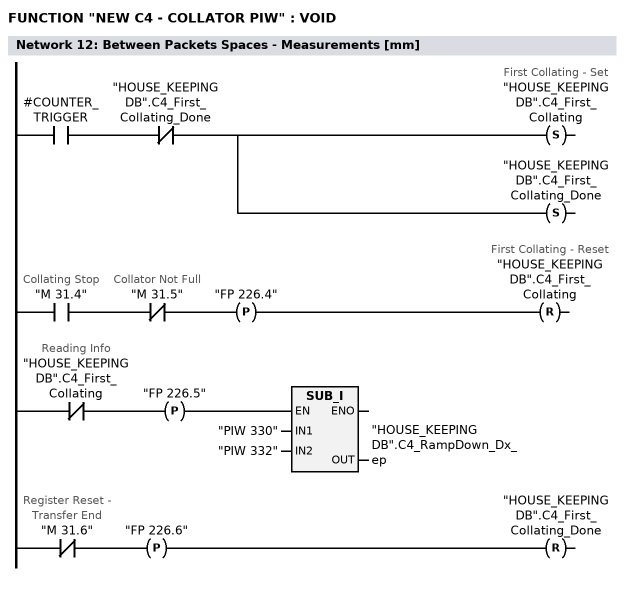

      A     #COUNTER_TRIGGER;
      AN    "HOUSE_KEEPING DB".C4_First_Collating_Done;
      S     "HOUSE_KEEPING DB".C4_First_Collating; // First Collating - Set
      S     "HOUSE_KEEPING DB".C4_First_Collating_Done;
//;
      A     "M 31.4"; // Collating Stop
      AN    "M 31.5"; // Collator Not Full
      FP    "FP 226.4";
      R     "HOUSE_KEEPING DB".C4_First_Collating; // First Collating - Reset
//;
      AN    "HOUSE_KEEPING DB".C4_First_Collating; // Reading Info
      FP    "FP 226.5";
      JCN   N1ST;

      L     "PIW 330"; // Direct Ch3 (was ACT_CNTV3, ~100 mS old)
      L     "PIW 332"; // Direct Ch2 (was ACT_CNTV2, ~100 mS old)
      -I    ;
      T     "HOUSE_KEEPING DB".C4_RampDown_Dx_ep;

N1ST: NOP   0;

      AN    "M 31.6"; // Register Reset - Transfer End
      FP    "FP 226.6";
      R     "HOUSE_KEEPING DB".C4_First_Collating_Done;
NETWORK
TITLE =Conveyor 4 - Surface Length Left (PulseUnit) - Measurements

      A     "M 31.1";
      S     "M 166.3";
//;
      A     "M 166.3";
      AN    "M 31.7";
      =     "FM350 DB".CONTROL_SIGNALS.SW_GATE3;
//;
      A     "M 166.3";
      A     "M 31.1";
      JNB   M663;
      L     "COLLATORS DB".Surface_Length_C4;
      L     "PIW 330"; // Direct Ch3 (was ACT_CNTV3, ~100 mS old)
      -D    ;
      T     "COLLATORS DB".Surface_Left_C4;
      L     0;
      >=I   ;
      JNB   T004;
      L     "COLLATORS DB".Surface_Left_C4;
      T     "COLLATORS DB".Surface_Length_Left_C4;

T004: CLR   ;

M663: CLR   ;
NETWORK
TITLE =Conveyor 4 - Space Between - Calculator

      A     "M 167.1";
      FP    "FP 154.2";
      JNB   M581;
      L     "COLLATORS DB".Surface_Left_C4;
      L     "COLLATORS DB".Frac_Packet_Length_C4;
      -I    ;
      T     "MW 214";

M581: CLR   ;

      A     "M 167.1";
      JNB   M671;
      A(    ;
      L     "COLLATORS DB".Surface_Left_C4;
      L     "MW 214";
      <=I   ;
      )     ;
      R     "M 167.1";

M671: CLR   ;
NETWORK
TITLE =Conveyor 4 - Collating Length Manager

      A     "M 166.3";
      AN    "M 30.4";
      A     "M 31.4";
      JNB   M304;
      L     "COLLATORS DB".Surface_Left_C4;
      L     "COLLATORS DB".Packet_Length_Frac_C4;
      <I    ;
      S     "M 30.4";

M304: CLR   ;

      A     "M 10.1";
      FP    "FP 154.7";
      O     "M 31.7";
      R     "M 30.4";
NETWORK
TITLE =Packet Length to HMI + Hysteresis

      A     "M 167.4";
      JNB   C167;
      A(    ;
      A(    ;
      L     "MW 202";
      L     "MW 204";
      >I    ;
      )     ;
      O     ;
      A(    ;
      L     "MW 202";
      L     "MW 206";
      <I    ;
      )     ;
      )     ;
      JNB   BYP5;
      L     "MW 202";
      T     "HMI_DB".WORD_PACKET_LENGTH;

BYP5: CLR   ;

      L     "MW 202";
      L     3.000000e+000;
      *R    ;
      L     1.000000e+002;
      /R    ;
      T     #R_TUBE_PERCENT;
      TRUNC ;
      T     #W_TUBE_PERCENT;
//;
      L     #W_TUBE_PERCENT;
      L     "MW 202";
      +I    ;
      T     "MW 204";
//;
      L     #W_TUBE_PERCENT;
      L     "MW 202";
      -I    ;
      T     "MW 206";
//;
      CLR   ;
      =     "M 167.4";

C167: CLR   ;
NETWORK
TITLE =Collator
//Collator House Keeping


NETWORK
TITLE =Collator Conveyor 4 - Clearing
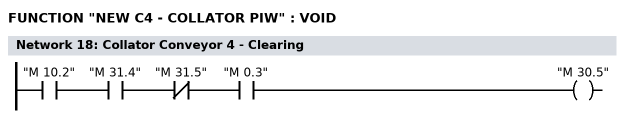

      A     "M 10.2";
      A     "M 31.4";
      AN    "M 31.5";
      A     "M 0.3";
      =     "M 30.5";
NETWORK
TITLE =Soft Timer 33 Reset - Clearing TimeOut 20s + Freeze Option

      A     "M 30.5";
      A     "A 44.3";
      A     "M 0.3";
      JCN   R331;
      JU    E331;

R331: L     L#0;
      T     "DB UTILITY".T33_ET;
      R     "DB UTILITY".T33_DN;

E331: NOP   0;
NETWORK
TITLE =Soft Timer 33 Add

      A     "M 30.5";
      A     "A 44.3";
      A     "M 0.3";
      AN    "DB UTILITY".Freeze_Sequence_2;
      AN    "DB UTILITY".T33_DN;
      JCN   E332;

      L     "DB UTILITY".T33_ET;
      L     "DB UTILITY".Scan_Cycle_Previous;
      ITD   ;
      +D    ;
      T     "DB UTILITY".T33_ET;

E332: NOP   0;
NETWORK
TITLE =Soft Timer 33 Done 20s

      L     "DB UTILITY".T33_ET;
      L     L#20000;
      >=D   ;
      =     "DB UTILITY".T33_DN;
NETWORK
TITLE =Collator Conveyor 4 - Clearing Surface - Run 2K Encoder Counts

      A     "M 30.5";
      A     "A 44.3";
      A     "M 0.3";
      JNB   M305;
      A(    ;
      L     "PIW 332"; // Direct Ch2 (was ACT_CNTV2, ~100 mS old)
      L     2000;
      >I    ;
      )     ;
      =     "M 30.3";

M305: CLR   ;
NETWORK
TITLE =Collator Conveyor 4 - Packet at the End !
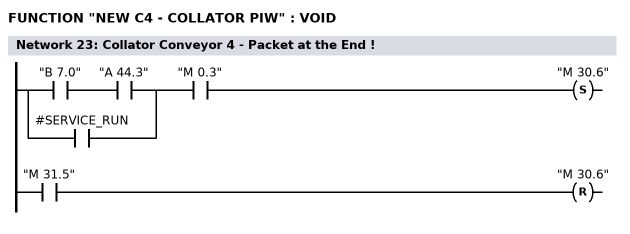

      A     "B 7.0";
      A     "A 44.3";
      O     #SERVICE_RUN;
      A     "M 0.3";
      S     "M 30.6";
//;
      A     "M 31.5";
      R     "M 30.6";
NETWORK
TITLE =Soft Timer 31 Reset - InFeed TimeOut 5s With Freeze Option

      A     "M 31.2";
      AN    "M 31.4";
      A     "A 44.3";
      A     "M 0.3";
      JCN   R311;
      JU    E311;

R311: L     L#0;
      T     "DB UTILITY".T31_ET;
      R     "DB UTILITY".T31_DN;

E311: NOP   0;
NETWORK
TITLE =Soft Timer 31 Add

      A     "M 31.2";
      AN    "M 31.4";
      A     "A 44.3";
      A     "M 0.3";
      AN    "DB UTILITY".Freeze_Sequence_2;
      AN    "DB UTILITY".T31_DN;
      JCN   E312;

      L     "DB UTILITY".T31_ET;
      L     "DB UTILITY".Scan_Cycle_Previous;
      ITD   ;
      +D    ;
      T     "DB UTILITY".T31_ET;

E312: NOP   0;
NETWORK
TITLE =Soft Timer 31 Done 5s
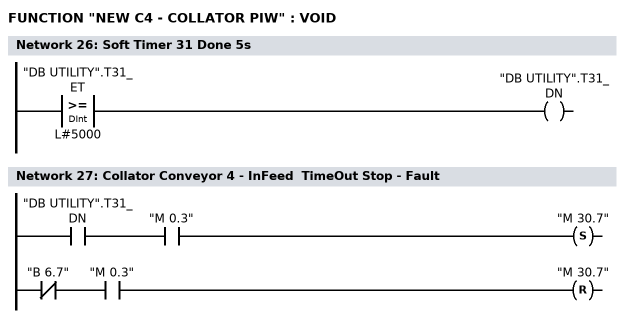

      L     "DB UTILITY".T31_ET;
      L     L#5000;
      >=D   ;
      =     "DB UTILITY".T31_DN;
NETWORK
TITLE =Collator Conveyor 4 - InFeed  TimeOut Stop - Fault

      A     "DB UTILITY".T31_DN;
      A     "M 0.3";
      S     "M 30.7";
//;
      AN    "B 6.7";
      A     "M 0.3";
      R     "M 30.7";
NETWORK
TITLE =Collator
//Collator Steps


NETWORK
TITLE =Collator Conveyor 4 - Steps Register - Reset

      A(    ;
      O     "M 31.7";
      O     "DB UTILITY".T33_DN;
      O     #INITIALISATION;
      O     "DB UTILITY".Conveyor_4_Disable;
      )     ;
      A     "M 0.3";
      JNB   INIT;
      L     W#16#0;
      T     "MW 31";
      S     "M 167.0";

INIT: CLR   ;
NETWORK
TITLE =Step 5N1  - Power ON
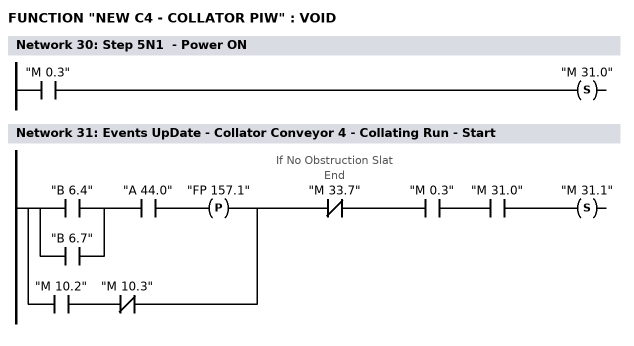

      A     "M 0.3";
      S     "M 31.0";
NETWORK
TITLE =Events UpDate - Collator Conveyor 4 - Collating Run - Start

      A(    ;
      A(    ;
      O     "B 6.4";
      O     "B 6.7";
      )     ;
      A     "A 44.0";
      FP    "FP 157.1";
      O     ;
      A     "M 10.2";
      AN    "M 10.3";
      )     ;
      AN    "M 33.7"; // If No Obstruction Slat End
      A     "M 0.3";
      A     "M 31.0";
      S     "M 31.1";
NETWORK
TITLE =Soft Timer 29 Reset - LB Obstruction Alarm 10s + Freeze Option

      A(    ;
      O     "B 6.4";
      O     "B 6.7";
      )     ;
      AN    "A 44.0";
      JCN   R281;
      JU    E281;

R281: L     L#0;
      T     "DB UTILITY".T29_ET;
      R     "DB UTILITY".T29_DN;

E281: NOP   0;
NETWORK
TITLE =Soft Timer 29 Add

      A(    ;
      O     "B 6.4";
      O     "B 6.7";
      )     ;
      AN    "A 44.0";
      AN    "DB UTILITY".Freeze_Sequence_2;
      AN    "DB UTILITY".T29_DN;
      JCN   E282;

      L     "DB UTILITY".T29_ET;
      L     "DB UTILITY".Scan_Cycle_Previous;
      ITD   ;
      +D    ;
      T     "DB UTILITY".T29_ET;

E282: NOP   0;
NETWORK
TITLE =Soft Timer 29 Done 10s
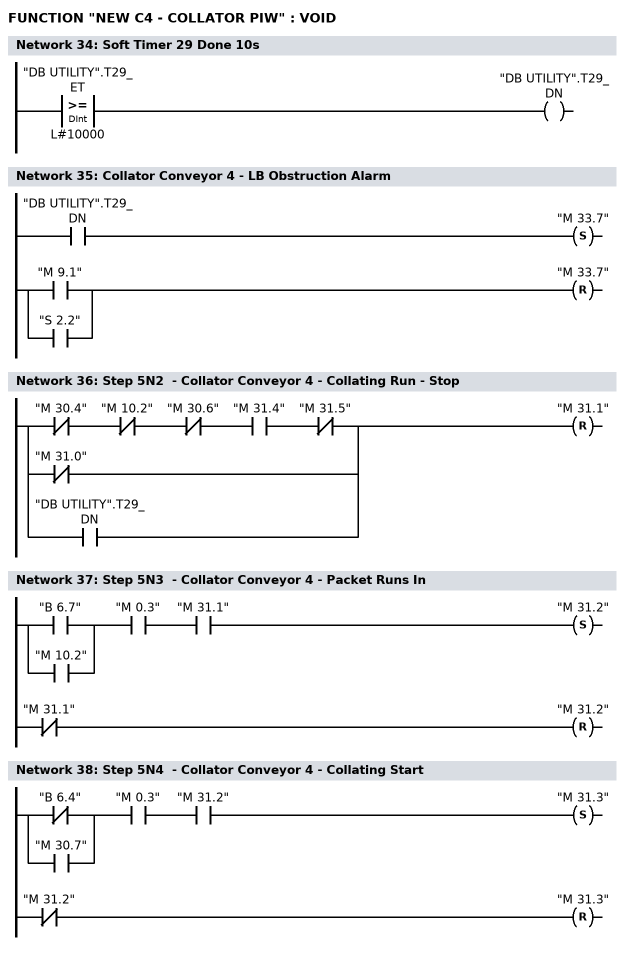

      L     "DB UTILITY".T29_ET;
      L     L#10000;
      >=D   ;
      =     "DB UTILITY".T29_DN;
NETWORK
TITLE =Collator Conveyor 4 - LB Obstruction Alarm

      A     "DB UTILITY".T29_DN;
      S     "M 33.7";
//;
      A(    ;
      O     "M 9.1";
      O     "S 2.2";
      )     ;
      R     "M 33.7";
NETWORK
TITLE =Step 5N2  - Collator Conveyor 4 - Collating Run - Stop

      A(    ;
      AN    "M 30.4";
      AN    "M 10.2";
      AN    "M 30.6";
      A     "M 31.4";
      AN    "M 31.5";
      ON    "M 31.0";
      O     "DB UTILITY".T29_DN;
      )     ;
      R     "M 31.1";
NETWORK
TITLE =Step 5N3  - Collator Conveyor 4 - Packet Runs In

      A(    ;
      O     "B 6.7";
      O     "M 10.2";
      )     ;
      A     "M 0.3";
      A     "M 31.1";
      S     "M 31.2";
//;
      AN    "M 31.1";
      R     "M 31.2";
NETWORK
TITLE =Step 5N4  - Collator Conveyor 4 - Collating Start

      A(    ;
      ON    "B 6.4";
      O     "M 30.7";
      )     ;
      A     "M 0.3";
      A     "M 31.2";
      S     "M 31.3";
//;
      AN    "M 31.2";
      R     "M 31.3";
NETWORK
TITLE =Step 5N5  - Collator Conveyor 4 - Collating Stop

      A(    ;
      AN    "B 6.7";
      AN(   ;
      AN    "M 10.2";
      A     "M 167.1";
      )     ;
      O     "M 30.7";
      )     ;
      A     "M 0.3";
      A     "M 31.3";
      S     "M 31.4";
//;
      AN    "M 31.3";
      R     "M 31.4";
NETWORK
TITLE =Step 5N6  - Collator Conveyor 4 - Full - Start Transfer
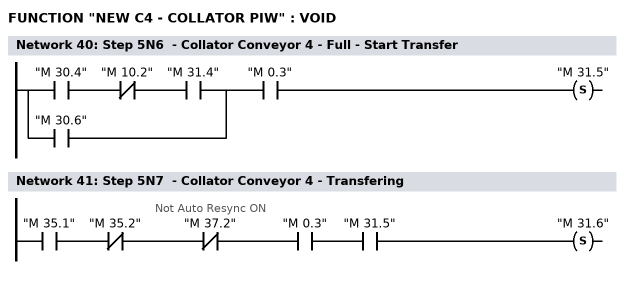

      A(    ;
      A     "M 30.4";
      AN    "M 10.2";
      A     "M 31.4";
      O     "M 30.6";
      )     ;
      A     "M 0.3";
      S     "M 31.5";
NETWORK
TITLE =Step 5N7  - Collator Conveyor 4 - Transfering

      A     "M 35.1";
      AN    "M 35.2";
      AN    "M 37.2"; // Not Auto Resync ON
      A     "M 0.3";
      A     "M 31.5";
      S     "M 31.6";
NETWORK
TITLE =Soft Timer 32 Reset - Transfer TimeOut 20s + Freeze Option

      A     "M 31.6";
      AN    "M 31.7";
      A     "A 44.3";
      A     "M 0.3";
      JCN   R321;
      JU    E321;

R321: L     L#0;
      T     "DB UTILITY".T32_ET;
      R     "DB UTILITY".T32_DN;

E321: NOP   0;
NETWORK
TITLE =Soft Timer 32 Add

      A     "M 31.6";
      AN    "M 31.7";
      A     "A 44.3";
      A     "M 0.3";
      AN    "DB UTILITY".Freeze_Sequence_2;
      AN    "DB UTILITY".T32_DN;
      JCN   E322;

      L     "DB UTILITY".T32_ET;
      L     "DB UTILITY".Scan_Cycle_Previous;
      ITD   ;
      +D    ;
      T     "DB UTILITY".T32_ET;

E322: NOP   0;
NETWORK
TITLE =Soft Timer 32 Done 20s
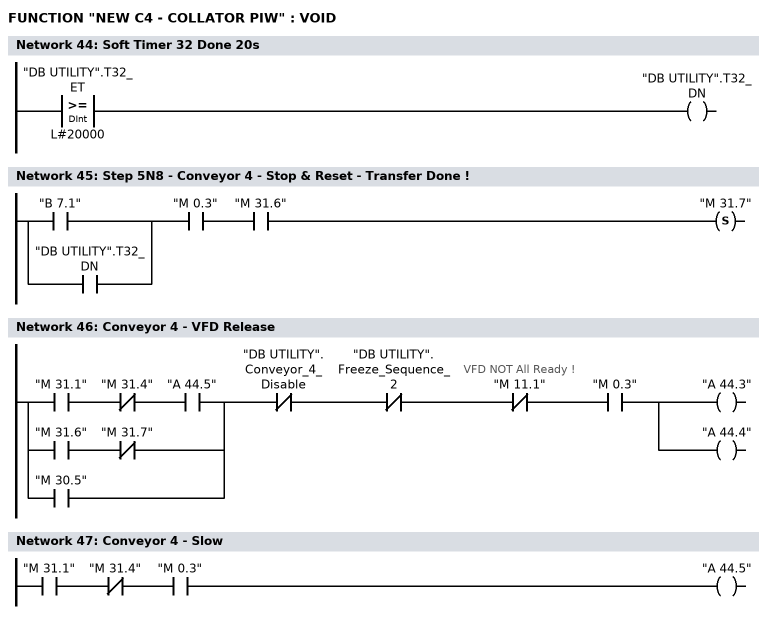

      L     "DB UTILITY".T32_ET;
      L     L#20000;
      >=D   ;
      =     "DB UTILITY".T32_DN;
NETWORK
TITLE =Step 5N8 - Conveyor 4 - Stop & Reset - Transfer Done !

      A(    ;
      O     "B 7.1";
      O     "DB UTILITY".T32_DN;
      )     ;
      A     "M 0.3";
      A     "M 31.6";
      S     "M 31.7";
NETWORK
TITLE =Conveyor 4 - VFD Release

      A(    ;
      A     "M 31.1";
      AN    "M 31.4";
      A     "A 44.5";
      O     ;
      A     "M 31.6";
      AN    "M 31.7";
      O     "M 30.5";
      )     ;
      AN    "DB UTILITY".Conveyor_4_Disable;
      AN    "DB UTILITY".Freeze_Sequence_2;
      AN    "M 11.1"; // VFD NOT All Ready !
      A     "M 0.3";
      =     "A 44.3";
      =     "A 44.4";
NETWORK
TITLE =Conveyor 4 - Slow

      A     "M 31.1";
      AN    "M 31.4";
      A     "M 0.3";
      =     "A 44.5";
END_FUNCTION

FUNCTION "NEW C5 - LINK" : VOID
TITLE =NEW FC934 (was FC1034) - Conveyor 5 - Link Pos.7
//Using "Soft Timer" cause S5T Timer cannot Pause/Freeze !...
NAME : POS_7
VERSION : 0.0


VAR_TEMP
  MAIN_SERVICE_2_SW : BOOL ;
  SERVICE_RUN : BOOL ;
  INITIALISATION : BOOL ;
END_VAR
BEGIN
NETWORK
TITLE =Conveyor 5 - Service

      A     "HMI_DB".ALL_SERVICE_ENABLE_SW;
      A     "HMI_DB".CONVEYOR_5_SERVICE_SW;
      A     "HMI_DB".SERVICE_SW_2_STATUS;
      =     #MAIN_SERVICE_2_SW;
//;
      A     #MAIN_SERVICE_2_SW;
      O     "M 34.1";
      JNB   CON5;
//;
      A     "HMI_DB".HMI_CONVEYOR_5_TEST_SSW;
      AN    "A 44.3";
      =     #SERVICE_RUN;
      S     "DB UTILITY".Conveyor_4_Disable;
//;
      A     "HMI_DB".SERVICE_INIT_PB;
      =     #INITIALISATION;
//;
      AN    #MAIN_SERVICE_2_SW;
      R     "HMI_DB".HMI_CONVEYOR_5_TEST_SSW;
      R     "DB UTILITY".Conveyor_4_Disable;

CON5: R     #SERVICE_RUN;
      R     #INITIALISATION;
      FP    "FP 158.5";
      =     "M 34.1";

NETWORK
TITLE =Service Mode
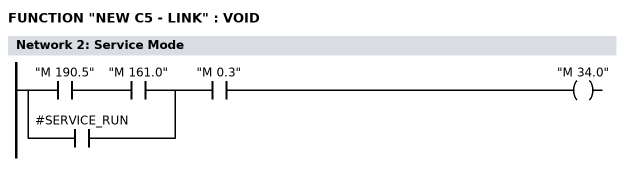

      A(    ;
      A     "M 190.5";
      A     "M 161.0";
      O     ;
      A     #SERVICE_RUN;
      )     ;
      A     "M 0.3";
      =     "M 34.0";

NETWORK
TITLE =Conveyor 5 - Steps Register - Reset

      A(    ;
      A     "M 35.1";
      AN    "M 35.2";
      A     "DB UTILITY".T35_DN;
      O     "M 35.4";
      O     #INITIALISATION;
      O     "DB UTILITY".Conveyor_5_Disable;
      )     ;
      A     "M 0.3";
      JC    M001;
      JU    M002;

M001: L     W#16#0;
      T     "MW 35";
      T     "HMI DB NEW".CONV_5_COUNT;

M002: NOP   0;

NETWORK
TITLE =Step 6N1 - Power ON
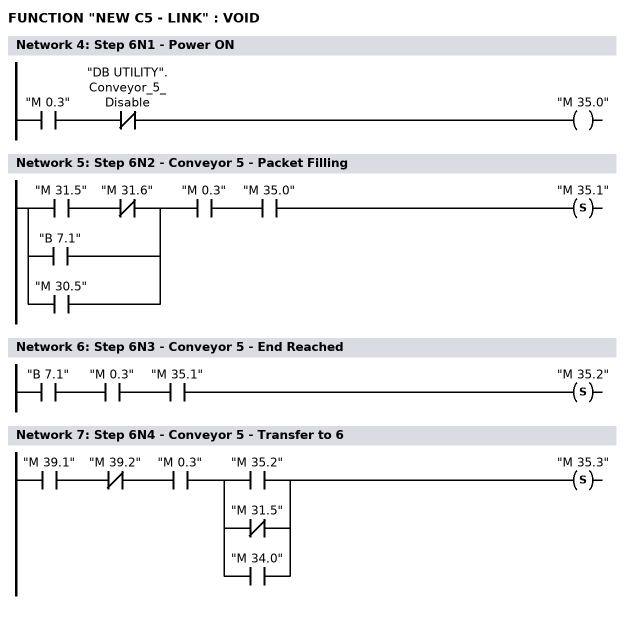

      A     "M 0.3";
      AN    "DB UTILITY".Conveyor_5_Disable;
      =     "M 35.0";

NETWORK
TITLE =Step 6N2 - Conveyor 5 - Packet Filling

      A(    ;
      A     "M 31.5";
      AN    "M 31.6";
      O     "B 7.1";
      O     "M 30.5";
      )     ;
      A     "M 0.3";
      A     "M 35.0";
      S     "M 35.1";

NETWORK
TITLE =Step 6N3 - Conveyor 5 - End Reached

      A     "B 7.1";
      A     "M 0.3";
      A     "M 35.1";
      S     "M 35.2";

NETWORK
TITLE =Step 6N4 - Conveyor 5 - Transfer to 6

      A     "M 39.1";
      AN    "M 39.2";
      A     "M 0.3";
      A(    ;
      O     "M 35.2";
      ON    "M 31.5";
      O     "M 34.0";
      )     ;
      S     "M 35.3";

NETWORK
TITLE =Soft Timer 35 Reset

      A(    ;
      A     "M 35.1";
      AN    "M 35.2";
      O     ;
      A     "M 35.3";
      AN    "M 35.4";
      A     "A 45.0";
      )     ;
      A     "M 0.3";
      JCN   R351;
      JU    E351;

R351: L     L#0;
      T     "DB UTILITY".T35_ET;
      R     "DB UTILITY".T35_DN;

E351: NOP   0;

NETWORK
TITLE =Soft Timer 35 Add

      A(    ;
      A     "M 35.1";
      AN    "M 35.2";
      O     ;
      A     "M 35.3";
      AN    "M 35.4";
      A     "A 45.0";
      )     ;
      A     "M 0.3";
      JCN   E352;
//;
      A     "DB UTILITY".Freeze_Sequence_2;
      A     "M 35.1";
      AN    "M 35.2";
      JC    E352;
//;
      AN    "DB UTILITY".T35_DN;
      JCN   E352;
//;
      L     "DB UTILITY".T35_ET;
      L     "DB UTILITY".Scan_Cycle_Previous;
      ITD   ;
      +D    ;
      T     "DB UTILITY".T35_ET;

E352: NOP   0;

NETWORK
TITLE =Soft Timer 35 Done 30s

      L     "DB UTILITY".T35_ET;
      L     L#30000; // [mS]
      >=D   ;
      =     "DB UTILITY".T35_DN;

NETWORK
TITLE =Automatic Re-Synchronization
//In Order to keep Synchronized,
//if Every Conditions are there, Conveyor 5 will do a Synchro Run 13sec after
//every 5 runs !
      A     "A 45.0"; // Count runs
      FP    "FP 169.7";
      JNB   ARS1;

      L     "MW 220"; // Count up
      L     1;
      +I    ;
      T     "MW 220";
//;
      L     10;
      >=I   ;
      JNB   ARS1;
//;
      S     "M 37.3"; // ARM after 5 runs
      L     0;
      T     "MW 220";

ARS1: NOP   0;

      A     "M 37.3"; // ARMED
      AN    "M 37.2"; // NOT already running
      AN    "DB UTILITY".Freeze_Sequence_2;
      AN    "A 45.0"; // wait end of run
      A     "M 35.0"; // power ON
      AN    "M 35.4"; // not in reset/stop
      JNB   ARS2;
//;
      L     "HMI_DB".CONV_4_COUNT; // Conveyor 4 Must be <= 2
      L     3;
      <I    ;
      JNB   ARS2;
//;
      L     "HMI_DB".CONV_5_COUNT;
      L     0; // Conveyor 5 Must NOT be Empty
      >I    ;
      JNB   ARS2;
//;
      L     "HMI_DB".CONV_6_COUNT;
      L     0; // Conveyor 6 Must be Empty
      ==I   ;
      JNB   ARS2;
//;
      AN    "B 7.2"; // Conveyor 6 Must be Empty
      AN    "M 10.0"; // Not Clearing
      JNB   ARS2;
//;
      S     "M 37.2"; // START 13s RUN
      R     "M 37.3"; // DISARM

ARS2: NOP   0;

      A     "M 37.2"; // Re-Sync ON
      L     S5T#13S;
      SD    "Timer 64";
//;
      A     "Timer 64"; // End Re-Sync if TimeOut 13s
      O     "B 7.1"; // or if Packet at END Sensor
      R     "M 37.2"; // Re-Sync OFF
NETWORK
TITLE =Automatic Re-Synchronization - Arm Timeout
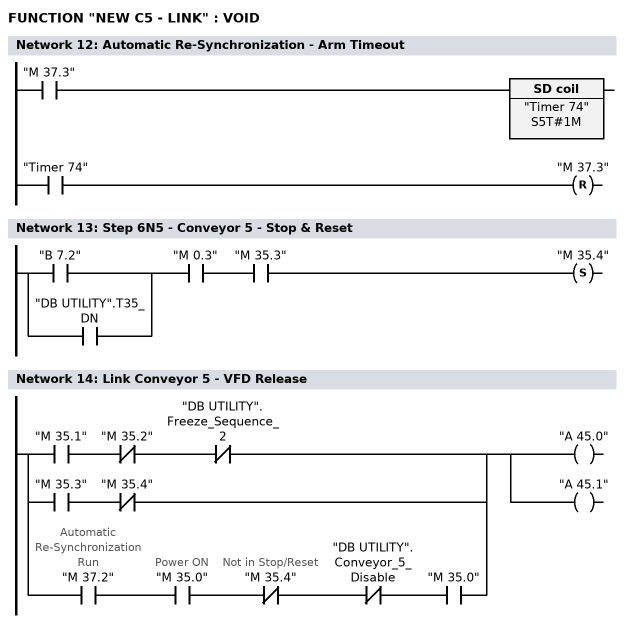

      A     "M 37.3";
      L     S5T#1M;
      SD    "Timer 74";
//;
      A     "Timer 74";
      R     "M 37.3";
NETWORK
TITLE =Step 6N5 - Conveyor 5 - Stop & Reset

      A(    ;
      O     "B 7.2";
      O     "DB UTILITY".T35_DN;
      )     ;
      A     "M 0.3";
      A     "M 35.3";
      S     "M 35.4";

NETWORK
TITLE =Link Conveyor 5 - VFD Release

      A(    ;
      A(    ;
      A     "M 35.1";
      AN    "M 35.2";
      AN    "DB UTILITY".Freeze_Sequence_2;
      )     ;
      O     ;
      A     "M 35.3";
      AN    "M 35.4";
      )     ;
      O     ;
      A(    ;
      A     "M 37.2"; // Automatic Re-Synchronization Run
      A     "M 35.0"; // Power ON
      AN    "M 35.4"; // Not in Stop/Reset
      )     ;
      AN    "DB UTILITY".Conveyor_5_Disable;
      A     "M 35.0";
      =     "A 45.0";
      =     "A 45.1";
END_FUNCTION

FUNCTION "NEW C6 - FLIP DELIV." : VOID
TITLE =NEW FC938 (was FC1038) - Conveyor 6 - Delivery to Flipper Pos.8
NAME : POS_8
VERSION : 0.0


VAR_TEMP
  MAIN_SERVICE_2_SW : BOOL ;
  SERVICE_RUN : BOOL ;
  INITIALISATION : BOOL ;
END_VAR
BEGIN
NETWORK
TITLE =Slat Conveyor - Service

      A     "HMI_DB".ALL_SERVICE_ENABLE_SW;
      A     "HMI_DB".CONVEYOR_6_SERVICE_SW;
      A     "HMI_DB".SERVICE_SW_2_STATUS;
      =     #MAIN_SERVICE_2_SW;
      CLR   ; // Fix: #INITIALISATION was never written
      =     #INITIALISATION;
//;
      A     #MAIN_SERVICE_2_SW;
      O     "M 38.1";
      JNB   CON6;
      A     "HMI_DB".HMI_CONVEYOR_6_TEST_SSW;
      =     #SERVICE_RUN;
      S     "DB UTILITY".Conveyor_5_Disable;
//;
      AN    #MAIN_SERVICE_2_SW;
      R     "HMI_DB".HMI_CONVEYOR_6_TEST_SSW;
      R     "DB UTILITY".Conveyor_5_Disable;

CON6: R     #SERVICE_RUN;
      R     #INITIALISATION;
      FP    "FP 158.6";
      =     "M 38.1";
NETWORK
TITLE =Flipper Delivery Conveyor 6 - Running TimeOut  30s
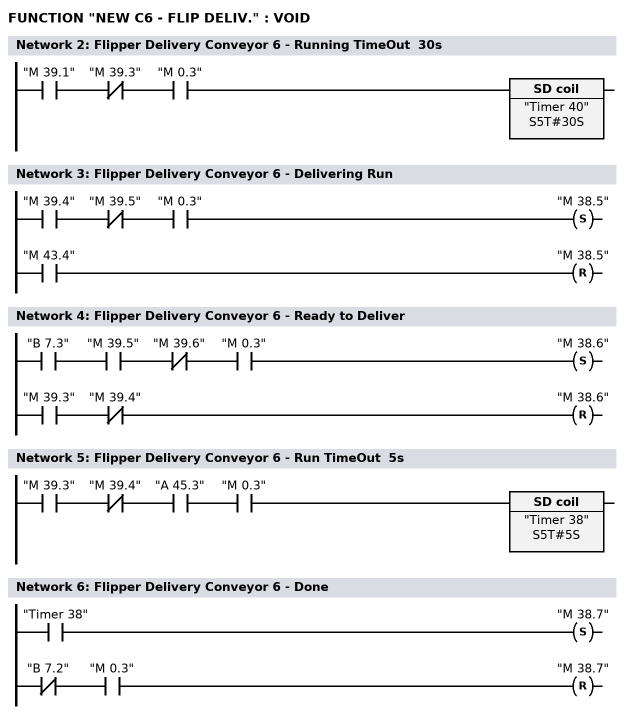

      A     "M 39.1";
      AN    "M 39.3";
      A     "M 0.3";
      L     S5T#30S;
      SD    "Timer 40";
NETWORK
TITLE =Flipper Delivery Conveyor 6 - Delivering Run

      A     "M 39.4";
      AN    "M 39.5";
      A     "M 0.3";
      S     "M 38.5";
//;
      A     "M 43.4";
      R     "M 38.5";
NETWORK
TITLE =Flipper Delivery Conveyor 6 - Ready to Deliver

      A     "B 7.3";
      A     "M 39.5";
      AN    "M 39.6";
      A     "M 0.3";
      S     "M 38.6";
//;
      A     "M 39.3";
      AN    "M 39.4";
      R     "M 38.6";
NETWORK
TITLE =Flipper Delivery Conveyor 6 - Run TimeOut  5s

      A     "M 39.3";
      AN    "M 39.4";
      A     "A 45.3";
      A     "M 0.3";
      L     S5T#5S;
      SD    "Timer 38";
NETWORK
TITLE =Flipper Delivery Conveyor 6 - Done

      A     "Timer 38";
      S     "M 38.7";
//;
      AN    "B 7.2";
      A     "M 0.3";
      R     "M 38.7";
NETWORK
TITLE =Conveyor 6 - Steps Register - Reset

      A(    ;
      O     "M 39.6";
      O     "Timer 40";
      O     #INITIALISATION;
      O     "DB UTILITY".Conveyor_6_Disable;
      )     ;
      A     "M 0.3";
      JC    M001;
      JU    M002;

M001: L     W#16#0;
      T     "MW 39";
      T     "MB 41";
      T     "HMI DB NEW".CONV_6_COUNT;

M002: NOP   0;
NETWORK
TITLE =Step 7N1 - Power ON
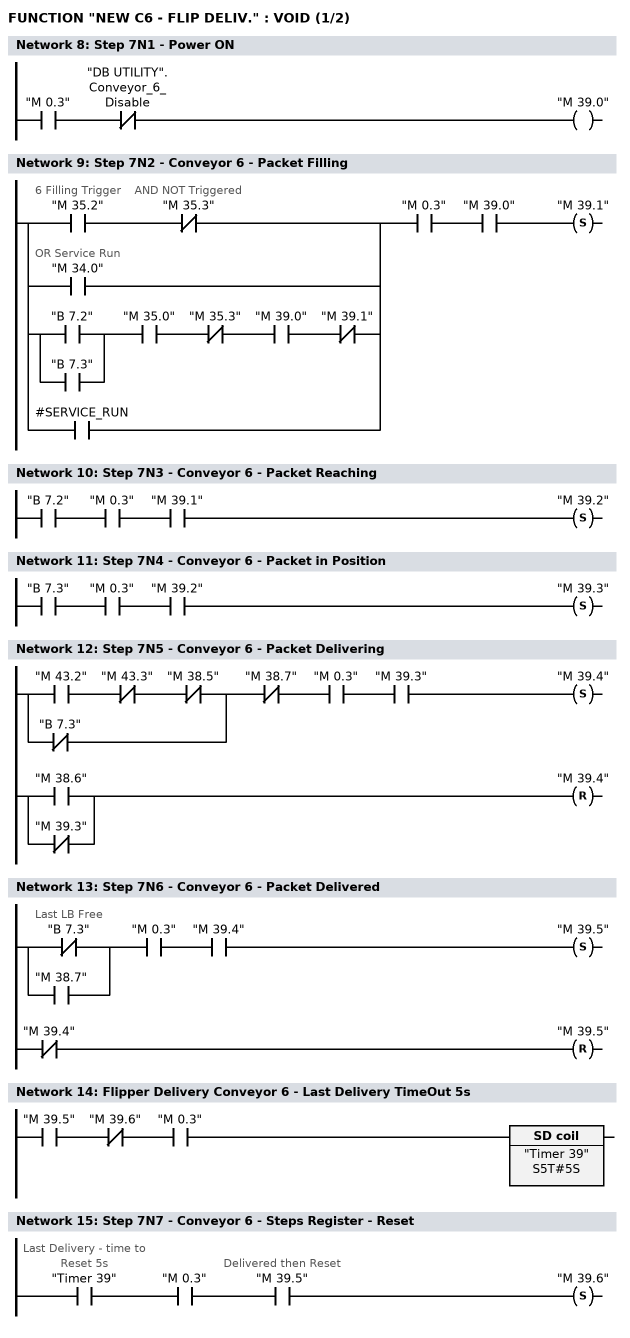

      A     "M 0.3";
      AN    "DB UTILITY".Conveyor_6_Disable;
      =     "M 39.0";
NETWORK
TITLE =Step 7N2 - Conveyor 6 - Packet Filling

      A(    ;

      A     "M 35.2"; // 6 Filling Trigger
      AN    "M 35.3"; // AND NOT Triggered
      O     "M 34.0"; // OR Service Run

      O     ;

      A(    ;
      O     "B 7.2";
      O     "B 7.3";
      )     ;
      A     "M 35.0";
      AN    "M 35.3";
      A     "M 39.0";
      AN    "M 39.1";

      O     ;

      A     #SERVICE_RUN;
      )     ;

      A     "M 0.3";
      A     "M 39.0";
      S     "M 39.1";
NETWORK
TITLE =Step 7N3 - Conveyor 6 - Packet Reaching

      A     "B 7.2";
      A     "M 0.3";
      A     "M 39.1";
      S     "M 39.2";
NETWORK
TITLE =Step 7N4 - Conveyor 6 - Packet in Position

      A     "B 7.3";
      A     "M 0.3";
      A     "M 39.2";
      S     "M 39.3";
NETWORK
TITLE =Step 7N5 - Conveyor 6 - Packet Delivering

      A(    ;
      A     "M 43.2";
      AN    "M 43.3";
      AN    "M 38.5";
      ON    "B 7.3";
      )     ;
      AN    "M 38.7";
      A     "M 0.3";
      A     "M 39.3";
      S     "M 39.4";
//;
      A(    ;
      O     "M 38.6";
      ON    "M 39.3";
      )     ;
      R     "M 39.4";
NETWORK
TITLE =Step 7N6 - Conveyor 6 - Packet Delivered

      A(    ;
      ON    "B 7.3"; // Last LB Free
      O     "M 38.7";
      )     ;
      A     "M 0.3";
      A     "M 39.4";
      S     "M 39.5";
//;
      AN    "M 39.4";
      R     "M 39.5";
NETWORK
TITLE =Flipper Delivery Conveyor 6 - Last Delivery TimeOut 5s

      A     "M 39.5";
      AN    "M 39.6";
      A     "M 0.3";
      L     S5T#5S;
      SD    "Timer 39";
NETWORK
TITLE =Step 7N7 - Conveyor 6 - Steps Register - Reset

      A     "Timer 39"; // Last Delivery - time to Reset 5s
      A     "M 0.3";
      A     "M 39.5"; // Delivered then Reset
      S     "M 39.6";
NETWORK
TITLE =Delivery Conveyor - VFD Release
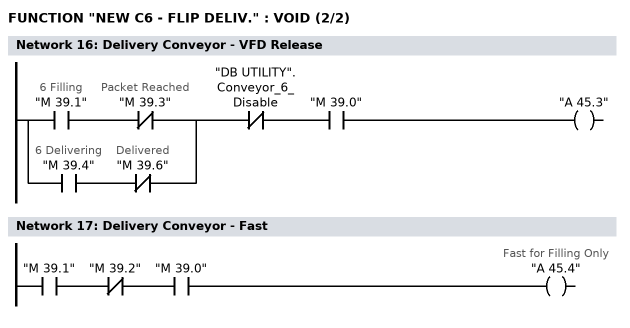

      A(    ;
      A     "M 39.1"; // 6 Filling
      AN    "M 39.3"; // Packet Reached
      O     ;
      A     "M 39.4"; // 6 Delivering
      AN    "M 39.6"; // Delivered
      )     ;
      AN    "DB UTILITY".Conveyor_6_Disable;
      A     "M 39.0";
      =     "A 45.3";
NETWORK
TITLE =Delivery Conveyor - Fast

      A     "M 39.1";
      AN    "M 39.2";
      A     "M 39.0";
      =     "A 45.4"; // Fast for Filling Only
END_FUNCTION

FUNCTION "NEW C7 - FLIPPER" : VOID
TITLE =NEW FC942 (was FC1042) - Flipper Pos.9
//Service : With FLIPPER Service SW "ON", To Flip, Hold the FLIP SW Until Reached
//or JOG to Position.
//v1.0 2026-11-23: Flipper conveyor stop time (Timer 42, step 8N5 -> 8N6) from
//DB15 "PACKET POSITION DB": one time per packet length class, set with the HMI
//arrows (FC1221, called here). Empty table = 1.5 s as before.
//v1.1 2026-11-24: calls FC1215 "PACKET POSITIONING" (was FC1221 "FLIPPER POS ADJ"),
//which also gives the C9 Pusher 2 stop time to FC950.
//v1.2 2026-11-24: DB15 symbol renamed "PACKET POSITION DB" - no code change.
NAME : POS_9
VERSION : 1.2


VAR_TEMP
  MAIN_SERVICE_2_SW : BOOL ;
  TIME_SW : BOOL ;
  FLIPPER_SERVICE_SW : BOOL ;
  FLIP : BOOL ;
  FLIP_CW : BOOL ;
  FLIP_CCW : BOOL ;
  CONVEYOR_7_RUN : BOOL ;
  INITIALISATION : BOOL ;
  POSITION_TIME : S5TIME ;
  T_ZOOLOO : TIME ;
  W_ZOOLOO_1 : WORD ;
  W_ZOOLOO_2 : WORD ;
END_VAR
BEGIN
NETWORK
TITLE =Stop Time per Packet Length - C7 + C9 (DB15, HMI Arrows)

      CALL "PACKET POSITIONING" ;

NETWORK
TITLE =Service Test

      A     "HMI_DB".ALL_SERVICE_ENABLE_SW;
      A     "HMI_DB".CONVEYOR_7_SERVICE_SW;
      A     "HMI_DB".SERVICE_SW_2_STATUS;
      R     "HMI_DB".SERVICE_SW_2_TIME_ADJ;
      =     #MAIN_SERVICE_2_SW;
//;
      A     #MAIN_SERVICE_2_SW;
      O     "M 42.3";
      JNB   FLIN;
      A     "HMI_DB".HMI_FLIPPER_SERVICE_SSW;
      =     #FLIPPER_SERVICE_SW;
      R     "HMI_DB".HMI_CONVEYOR_7_TEST_SSW;
//;
      A     "HMI_DB".HMI_CONVEYOR_7_TEST_SSW;
      =     #CONVEYOR_7_RUN;
      R     "HMI_DB".HMI_FLIPPER_SERVICE_SSW;
//;
      A     "HMI_DB".SERVICE_SW_2_TIME_ADJ;
      =     #TIME_SW;
//;
      AN    "P 8.0";
      S     "M 46.0";
      FP    "FP 168.5";
      S     "M 46.5";
//;
      AN    "P 8.1";
      R     "M 46.0";
      FP    "FP 168.6";
      S     "M 46.5";
//;
      A     #FLIPPER_SERVICE_SW;
      AN    "HMI_DB".HMI_FLIPPER_FLIP_SSW;
      L     S5T#3S;
      SE    "Timer 46";
//;
      A     "Timer 46";
      FN    "FN 155.1";
      R     "M 46.5";
//;
      A     #FLIPPER_SERVICE_SW;
      A     "HMI_DB".HMI_FLIPPER_FLIP_SSW;
      AN    "M 46.0";
      AN    "Timer 46";
      AN    "M 46.5";
      =     #FLIP_CW;
//;
      A     #FLIPPER_SERVICE_SW;
      A     "HMI_DB".HMI_FLIPPER_FLIP_SSW;
      A     "M 46.0";
      AN    "Timer 46";
      AN    "M 46.5";
      =     #FLIP_CCW;
//;
      A     "HMI_DB".HMI_CONVEYOR_7_TEST_SSW;
      =     #CONVEYOR_7_RUN;
//;
      A(    ;
      O     #FLIPPER_SERVICE_SW;
      O     #CONVEYOR_7_RUN;
      )     ;
      S     "DB UTILITY".Conveyor_6_Disable;
//;
      AN    #MAIN_SERVICE_2_SW;
      R     "HMI_DB".HMI_CONVEYOR_7_TEST_SSW;
      R     "HMI_DB".HMI_FLIPPER_SERVICE_SSW;
      R     "HMI_DB".HMI_FLIPPER_FLIP_SSW;
      R     "HMI_DB".SERVICE_SW_2_TIME_ADJ;
      R     "DB UTILITY".Conveyor_6_Disable;

FLIN: R     #TIME_SW;
      R     #FLIPPER_SERVICE_SW;
      R     #FLIP_CW;
      R     #FLIP_CCW;
      R     #CONVEYOR_7_RUN;
      FP    "FP 158.7";
      =     "M 42.3";
//;
      A     "HMI_DB".SERVICE_INIT_PB;
      A     #MAIN_SERVICE_2_SW;
      A     #FLIPPER_SERVICE_SW;
      =     #INITIALISATION;
NETWORK
TITLE =Flipper - Flip Status
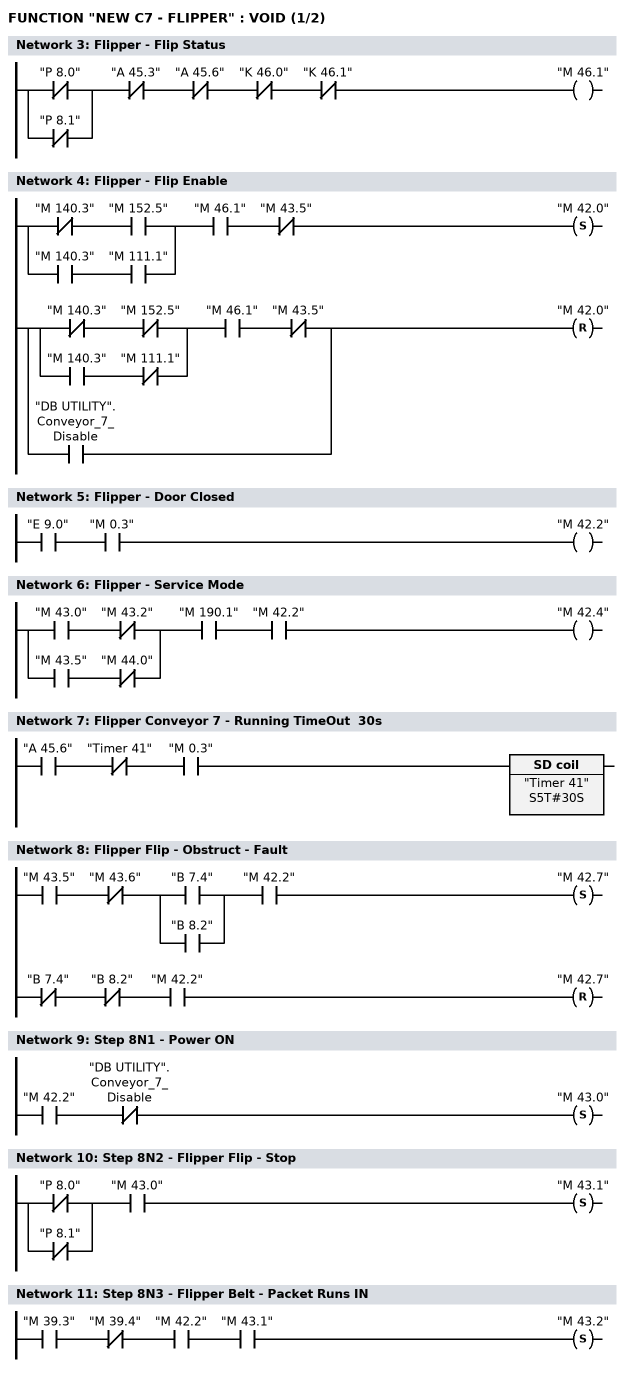

      A(    ;
      ON    "P 8.0";
      ON    "P 8.1";
      )     ;
      AN    "A 45.3";
      AN    "A 45.6";
      AN    "K 46.0";
      AN    "K 46.1";
      =     "M 46.1";
NETWORK
TITLE =Flipper - Flip Enable

      A(    ;
      AN    "M 140.3";
      A     "M 152.5";
      O     ;
      A     "M 140.3";
      A     "M 111.1";
      )     ;
      A     "M 46.1";
      AN    "M 43.5";
      S     "M 42.0";
//;
      A(    ;
      AN    "M 140.3";
      AN    "M 152.5";
      O     ;
      A     "M 140.3";
      AN    "M 111.1";
      )     ;
      A     "M 46.1";
      AN    "M 43.5";
      O     "DB UTILITY".Conveyor_7_Disable;
      R     "M 42.0";
NETWORK
TITLE =Flipper - Door Closed

      A     "E 9.0";
      A     "M 0.3";
      =     "M 42.2";
NETWORK
TITLE =Flipper - Service Mode

      A(    ;
      A     "M 43.0";
      AN    "M 43.2";
      O     ;
      A     "M 43.5";
      AN    "M 44.0";
      )     ;
      A     "M 190.1";
      A     "M 42.2";
      =     "M 42.4";
NETWORK
TITLE =Flipper Conveyor 7 - Running TimeOut  30s

      A     "A 45.6";
      AN    "Timer 41";
      A     "M 0.3";
      L     S5T#30S;
      SD    "Timer 41";
NETWORK
TITLE =Flipper Flip - Obstruct - Fault

      A     "M 43.5";
      AN    "M 43.6";
      A(    ;
      O     "B 7.4";
      O     "B 8.2";
      )     ;
      A     "M 42.2";
      S     "M 42.7";
//;
      AN    "B 7.4";
      AN    "B 8.2";
      A     "M 42.2";
      R     "M 42.7";
NETWORK
TITLE =Step 8N1 - Power ON

      A     "M 42.2";
      AN    "DB UTILITY".Conveyor_7_Disable;
      S     "M 43.0";
NETWORK
TITLE =Step 8N2 - Flipper Flip - Stop

      A(    ;
      ON    "P 8.0";
      ON    "P 8.1";
      )     ;
      A     "M 43.0";
      S     "M 43.1";
NETWORK
TITLE =Step 8N3 - Flipper Belt - Packet Runs IN

      A     "M 39.3";
      AN    "M 39.4";
      A     "M 42.2";
      A     "M 43.1";
      S     "M 43.2";
NETWORK
TITLE =Step 8N4 - Flipper Conveyor 7 - Packet Runs IN
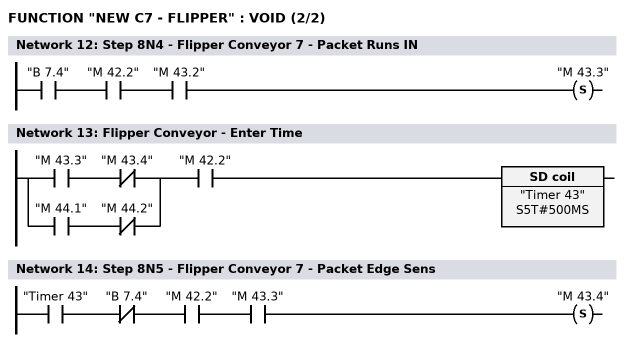

      A     "B 7.4";
      A     "M 42.2";
      A     "M 43.2";
      S     "M 43.3";
NETWORK
TITLE =Flipper Conveyor - Enter Time

      A(    ;
      A     "M 43.3";
      AN    "M 43.4";
      O     ;
      A     "M 44.1";
      AN    "M 44.2";
      )     ;
      A     "M 42.2";
      L     S5T#500MS;
      SD    "Timer 43";
NETWORK
TITLE =Step 8N5 - Flipper Conveyor 7 - Packet Edge Sens

      A     "Timer 43";
      AN    "B 7.4";
      A     "M 42.2";
      A     "M 43.3";
      S     "M 43.4";
NETWORK
TITLE =Time Convertion - Lateral Packet Position to Flipper - Adj.(HMI)
//   A     M    140.3
      AN    "M 6.7";
      FP    "FP 147.0";
      JNB   BYP1;
      L     "HMI_DB".CONV_7_POS_mS; // Integer contains MILLISECOND seconds
      L     50; // mS
      *I    ;
      T     #W_ZOOLOO_1;
      ITD   ;
      T     #T_ZOOLOO; // Double Int

      CALL "TIM_S5TI" (
           IN                       := #T_ZOOLOO,// Integer
           RET_VAL                  := #POSITION_TIME);// Simatic Time

      L     #POSITION_TIME;
      T     "MW 186"; // Simatic Time
//;
      L     #W_ZOOLOO_1;
      L     10;
      /I    ;
      T     #W_ZOOLOO_2;
//;
      A(    ;
      L     #W_ZOOLOO_2;
      L     "MW 192";
      <>I   ;
      )     ;
      JNB   BYP1;
      L     #W_ZOOLOO_2; // Simatic Time
      T     "HMI_DB".DELAY_DISPLAY_7;
      T     "MW 192";

BYP1: CLR   ;

      A     "M 140.3";
      A     "M 43.4";
      AN    "M 43.5";
      A     "M 42.2";
      A     "M 0.3";
      L     "MW 186"; // Simatic Time
      SD    "Timer 60";
NETWORK
TITLE =Flipper Conveyor Stop - Packet in Position
//     OPN   "DB LAUER"
//;
//      CALL  "LAUER TIME"
//       QUEL :=DBW242
//       _TIME:=MW122
//;
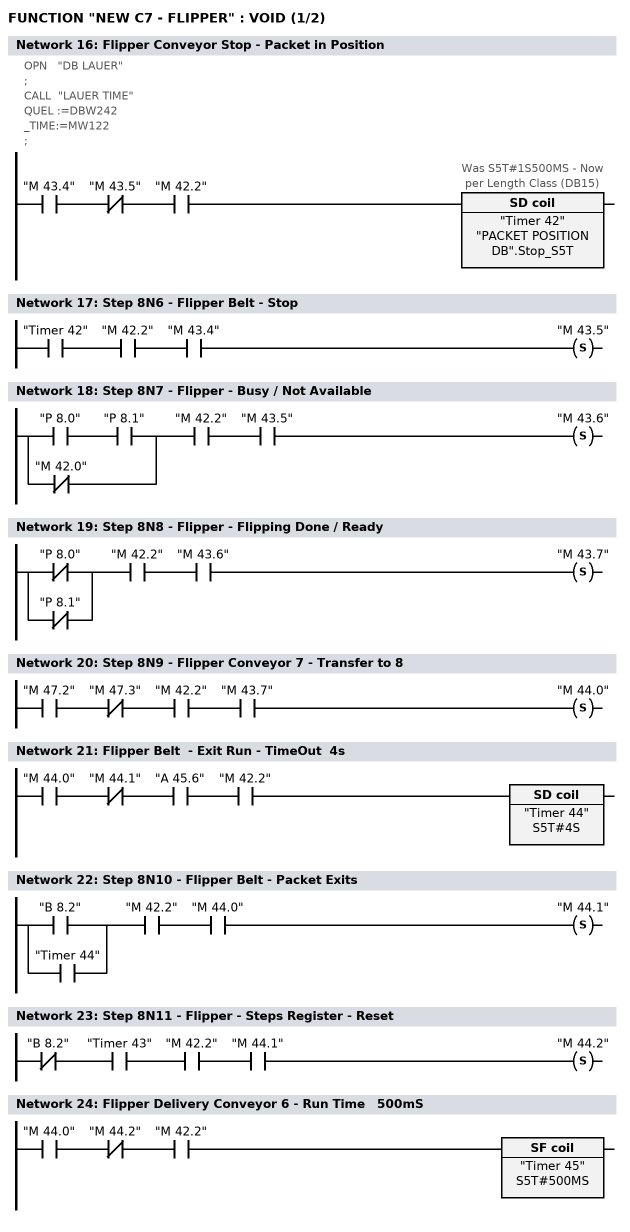
      A     "M 43.4";
      AN    "M 43.5";
      A     "M 42.2";
// L     MW   122
      L     "PACKET POSITION DB".Stop_S5T; // Was S5T#1S500MS - Now per Length Class (DB15)
      SD    "Timer 42";
NETWORK
TITLE =Step 8N6 - Flipper Belt - Stop

      A     "Timer 42";
//    O     T     60
      A     "M 42.2";
      A     "M 43.4";
      S     "M 43.5";
NETWORK
TITLE =Step 8N7 - Flipper - Busy / Not Available

      A(    ;
      A     "P 8.0";
      A     "P 8.1";
      ON    "M 42.0";
      )     ;
      A     "M 42.2";
      A     "M 43.5";
      S     "M 43.6";
NETWORK
TITLE =Step 8N8 - Flipper - Flipping Done / Ready

      A(    ;
      ON    "P 8.0";
      ON    "P 8.1";
      )     ;
      A     "M 42.2";
      A     "M 43.6";
      S     "M 43.7";
NETWORK
TITLE =Step 8N9 - Flipper Conveyor 7 - Transfer to 8

      A     "M 47.2";
      AN    "M 47.3";
      A     "M 42.2";
      A     "M 43.7";
      S     "M 44.0";
NETWORK
TITLE =Flipper Belt  - Exit Run - TimeOut  4s

      A     "M 44.0";
      AN    "M 44.1";
      A     "A 45.6";
      A     "M 42.2";
      L     S5T#4S;
      SD    "Timer 44";
NETWORK
TITLE =Step 8N10 - Flipper Belt - Packet Exits

      A(    ;
      O     "B 8.2";
      O     "Timer 44";
      )     ;
      A     "M 42.2";
      A     "M 44.0";
      S     "M 44.1";
NETWORK
TITLE =Step 8N11 - Flipper - Steps Register - Reset

      AN    "B 8.2";
      A     "Timer 43";
      A     "M 42.2";
      A     "M 44.1";
      S     "M 44.2";
NETWORK
TITLE =Flipper Delivery Conveyor 6 - Run Time   500mS

      A     "M 44.0";
      AN    "M 44.2";
      A     "M 42.2";
      L     S5T#500MS;
      SF    "Timer 45";
NETWORK
TITLE =Flipper Conveyor - VFD Release
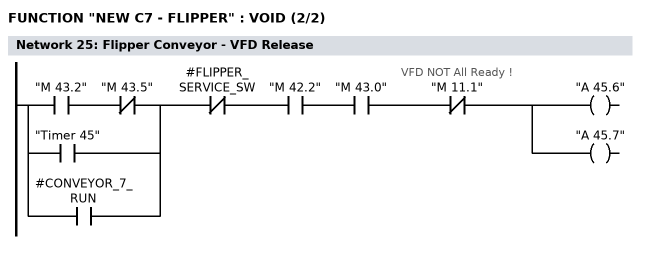

      A(    ;
      A     "M 43.2";
      AN    "M 43.5";
      O     "Timer 45";
      O     #CONVEYOR_7_RUN;
      )     ;
      AN    #FLIPPER_SERVICE_SW;
      A     "M 42.2";
      A     "M 43.0";
      AN    "M 11.1"; // VFD NOT All Ready !
      =     "A 45.6";
      =     "A 45.7";
NETWORK
TITLE =Flipper
//Flipper Action
NETWORK
TITLE =Flipper Flip - Steps Register - Reset

      A(    ;
      A     "M 190.1";
      A     "M 171.4";
      A     "M 171.5";
      O     "M 44.2";
      O     "Timer 41";
      O     #INITIALISATION;
      O     "DB UTILITY".Conveyor_7_Disable;
      )     ;
      A     "M 42.2";
      JC    M001;
      JU    M002;

M001: L     W#16#0;
      T     "MW 43";

M002: NOP   0;
NETWORK
TITLE =Events UpDate - Flipper Flip 1 - CW
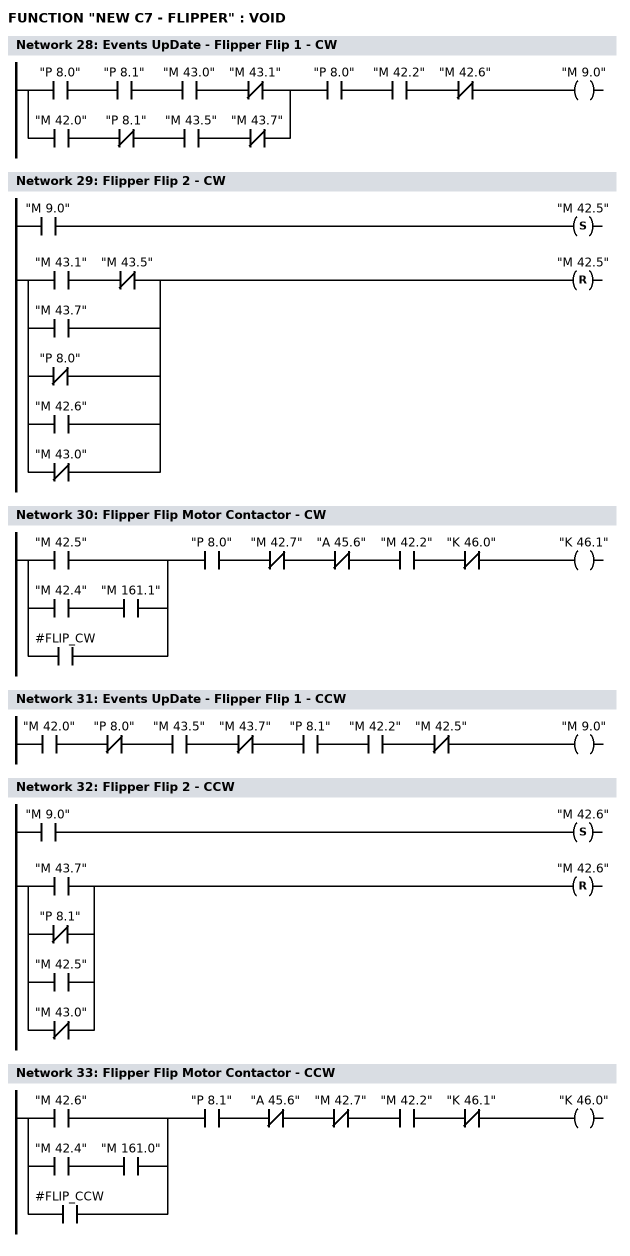

      A(    ;
      A     "P 8.0";
      A     "P 8.1";
      A     "M 43.0";
      AN    "M 43.1";
      O     ;
      A     "M 42.0";
      AN    "P 8.1";
      A     "M 43.5";
      AN    "M 43.7";
      )     ;
      A     "P 8.0";
      A     "M 42.2";
      AN    "M 42.6";
      =     "M 9.0";
NETWORK
TITLE =Flipper Flip 2 - CW

      A     "M 9.0";
      S     "M 42.5";
//;
      A(    ;
      A     "M 43.1";
      AN    "M 43.5";
      O     ;
      A     "M 43.7";
      O     ;
      AN    "P 8.0";
      O     "M 42.6";
      ON    "M 43.0";
      )     ;
      R     "M 42.5";
NETWORK
TITLE =Flipper Flip Motor Contactor - CW

      A(    ;
      A     "M 42.5";
      O     ;
      A     "M 42.4";
      A     "M 161.1";
      O     ;
      A     #FLIP_CW;
      )     ;
      A     "P 8.0";
      AN    "M 42.7";
      AN    "A 45.6";
      A     "M 42.2";
      AN    "K 46.0";
      =     "K 46.1";
NETWORK
TITLE =Events UpDate - Flipper Flip 1 - CCW

      A(    ;
      A     "M 42.0";
      AN    "P 8.0";
      A     "M 43.5";
      AN    "M 43.7";
      )     ;
      A     "P 8.1";
      A     "M 42.2";
      AN    "M 42.5";
      =     "M 9.0";
NETWORK
TITLE =Flipper Flip 2 - CCW

      A     "M 9.0";
      S     "M 42.6";
//;
      A(    ;
      A     "M 43.7";
      O     ;
      AN    "P 8.1";
      O     "M 42.5";
      ON    "M 43.0";
      )     ;
      R     "M 42.6";
NETWORK
TITLE =Flipper Flip Motor Contactor - CCW

      A(    ;
      A     "M 42.6";
      O     ;
      A     "M 42.4";
      A     "M 161.0";
      O     ;
      A     #FLIP_CCW;
      )     ;
      A     "P 8.1";
      AN    "A 45.6";
      AN    "M 42.7";
      A     "M 42.2";
      AN    "K 46.1";
      =     "K 46.0";
END_FUNCTION

FUNCTION "NEW C8 - TURNTABLE" : VOID
TITLE =NEW FC948 (was FC1048) - Turn Table Pos.10
//
NAME : POS_10
VERSION : 0.0


VAR_TEMP
  MAIN_SERVICE_2_SW : BOOL ;
  TURNTABLE_SERVICE_SW : BOOL ;
  CONVEYOR_SERVICE_SW : BOOL ;
  TURNTABLE_ROUNDTRIP : BOOL ;
  TURN_CW : BOOL ;
  TURN_CCW : BOOL ;
  AUTO_HOME_SERVICE : BOOL ;
  CONV_FWD : BOOL ;
  CONV_REV : BOOL ;
  INITIALISATION : BOOL ;
  ZOOLOO : TIME ;
  PACKET_LENGTH : REAL ;
  RUN_TIME : REAL ;
END_VAR
BEGIN
NETWORK
TITLE =Service Test

      A     "HMI_DB".ALL_SERVICE_ENABLE_SW;
      A     "HMI_DB".CONVEYOR_8_SERVICE_SW;
      A     "HMI_DB".SERVICE_SW_2_STATUS;
      =     #MAIN_SERVICE_2_SW;
//;
      A     #MAIN_SERVICE_2_SW;
      O     "M 46.7";
      JNB   TURN;
      A     "HMI_DB".HMI_CONVEYOR_8_TEST_SSW;
      =     #CONVEYOR_SERVICE_SW;
      R     "HMI_DB".TURNTABLE_SERVICE_SSW;
//;
      A     "HMI_DB".TURNTABLE_SERVICE_SSW;
      =     #TURNTABLE_SERVICE_SW;
      R     "HMI_DB".HMI_CONVEYOR_8_TEST_SSW;
//;
      A(    ;
      O     #CONVEYOR_SERVICE_SW;
      O     #TURNTABLE_SERVICE_SW;
      )     ;
      =     "HMI_DB".TURNTABLE_SERVICE_PBSHOW;
      S     "DB UTILITY".Conveyor_7_Disable;
//;
      A     "HMI_DB".TURNTABLE_RNDTRIP;
      S     "DB UTILITY".Conveyor_7_Disable;
//;
      A     "HMI_DB".SERVICE_INIT_PB;
      =     #AUTO_HOME_SERVICE;
//;
      A     #TURNTABLE_SERVICE_SW;
      A     "HMI_DB".HMI_TURNTABLE_CCW_SSW;
      AN    #TURN_CW;
      =     #TURN_CCW;
//;
      A     #TURNTABLE_SERVICE_SW;
      A     "HMI_DB".HMI_TURNTABLE_CW_SSW;
      AN    #TURN_CCW;
      =     #TURN_CW;
//;
      AN    #TURNTABLE_SERVICE_SW;
      =     "HMI_DB".RNDTRIP_PB_VISIBLE;
//;
      AN    #TURNTABLE_SERVICE_SW;
      A     "HMI_DB".TURNTABLE_RNDTRIP;
      =     #TURNTABLE_ROUNDTRIP;
//;
      A     #CONVEYOR_SERVICE_SW;
      A     "HMI_DB".HMI_TURNTABLE_CCW_SSW;
      AN    #CONV_FWD;
      =     #CONV_REV;
//;
      A     #CONVEYOR_SERVICE_SW;
      A     "HMI_DB".HMI_TURNTABLE_CW_SSW;
      AN    #CONV_REV;
      =     #CONV_FWD;
//;
      A     "HMI_DB".SERVICE_INIT_PB;
      A     #TURNTABLE_SERVICE_SW;
      =     #INITIALISATION;
//;
      AN    #MAIN_SERVICE_2_SW;
      R     "HMI_DB".TURNTABLE_SERVICE_SSW;
      R     "DB UTILITY".Conveyor_7_Disable;
      R     "HMI_DB".HMI_CONVEYOR_8_TEST_SSW;
      R     "HMI_DB".TURNTABLE_SERVICE_PBSHOW;
      R     "HMI_DB".HMI_TURNTABLE_CCW_SSW;
      R     "HMI_DB".HMI_TURNTABLE_CW_SSW;
      R     "HMI_DB".TURNTABLE_RNDTRIP;
      R     "HMI_DB".RNDTRIP_PB_VISIBLE;

TURN: R     #TURNTABLE_SERVICE_SW;
      R     #CONVEYOR_SERVICE_SW;
      R     #AUTO_HOME_SERVICE;
      R     #TURNTABLE_ROUNDTRIP;
      R     #INITIALISATION;
      R     #TURN_CW;
      R     #TURN_CCW;
      R     #CONV_FWD;
      R     #CONV_REV;
      FP    "FP 169.0";
      =     "M 46.7";
NETWORK
TITLE =Turn Direction - Turn Table Turn SW  1:CCW - 0:CW
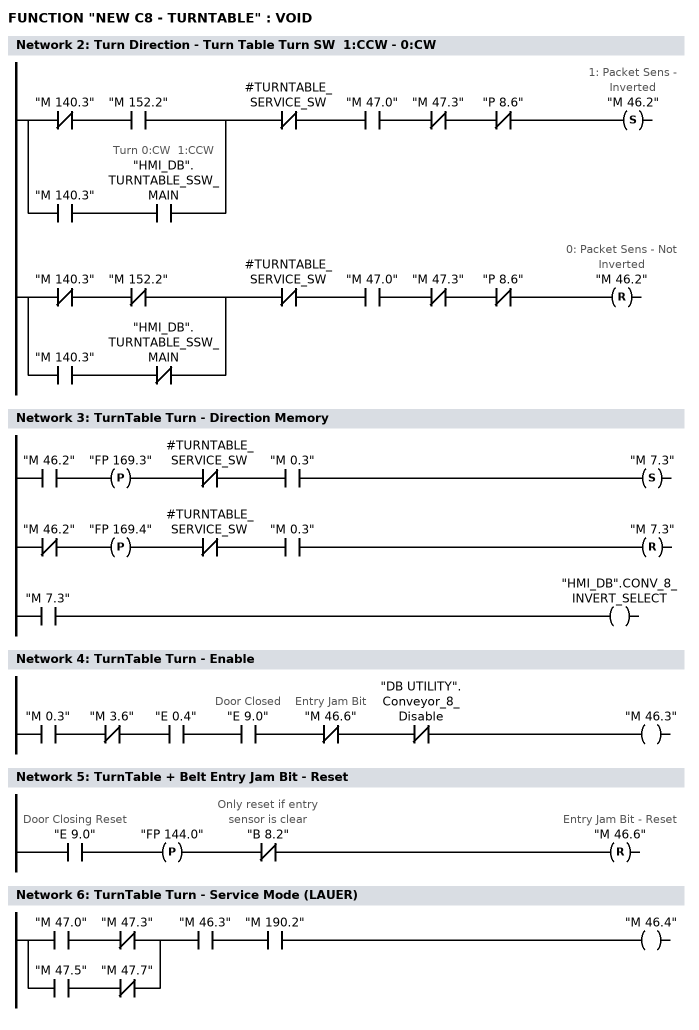

      A(    ;
      A(    ;
      AN    "M 140.3";
      A     "M 152.2";
      O     ;
      A     "M 140.3";
      A     "HMI_DB".TURNTABLE_SSW_MAIN; // Turn 0:CW  1:CCW
      )     ;
      AN    #TURNTABLE_SERVICE_SW;
      )     ;
      A     "M 47.0";
      AN    "M 47.3";
      AN    "P 8.6";
      S     "M 46.2"; // 1: Packet Sens - Inverted
//;
      A(    ;
      A(    ;
      AN    "M 140.3";
      AN    "M 152.2";
      O     ;
      A     "M 140.3";
      AN    "HMI_DB".TURNTABLE_SSW_MAIN;
      )     ;
      AN    #TURNTABLE_SERVICE_SW;
      )     ;
      A     "M 47.0";
      AN    "M 47.3";
      AN    "P 8.6";
      R     "M 46.2"; // 0: Packet Sens - Not Inverted
NETWORK
TITLE =TurnTable Turn - Direction Memory

      A     "M 46.2";
      FP    "FP 169.3";
      AN    #TURNTABLE_SERVICE_SW;
      A     "M 0.3";
      S     "M 7.3";
//;
      AN    "M 46.2";
      FP    "FP 169.4";
      AN    #TURNTABLE_SERVICE_SW;
      A     "M 0.3";
      R     "M 7.3";
//;
      A     "M 7.3";
      =     "HMI_DB".CONV_8_INVERT_SELECT;
NETWORK
TITLE =TurnTable Turn - Enable

      A     "M 0.3";
      AN    "M 3.6";
      A     "E 0.4";
      A     "E 9.0"; // Door Closed
      AN    "M 46.6"; // Entry Jam Bit
      AN    "DB UTILITY".Conveyor_8_Disable;
      =     "M 46.3";
NETWORK
TITLE =TurnTable + Belt Entry Jam Bit - Reset

      A     "E 9.0"; // Door Closing Reset
      FP    "FP 144.0";
      AN    "B 8.2"; // Only reset if entry sensor is clear
      R     "M 46.6"; // Entry Jam Bit - Reset
NETWORK
TITLE =TurnTable Turn - Service Mode (LAUER)

      A(    ;
      A     "M 47.0";
      AN    "M 47.3";
      O     ;
      A     "M 47.5";
      AN    "M 47.7";
      )     ;
      A     "M 46.3";
      A     "M 190.2";
      =     "M 46.4";
NETWORK
TITLE =Steps
//TurnTable Steps


NETWORK
TITLE =Step 9N0 - TurnTable Steps Register - Reset

      A(    ;
      A     "M 190.2";
      A     "M 171.4";
      A     "M 171.5";
      O     "M 48.4";
      O     #INITIALISATION;
      )     ;
      A     "M 46.3";
      O     "M 46.6"; // Entry Jam Fault - Reset
      JC    M001;
      JU    M002;

M001: L     W#16#0;
      T     "MW 47";

M002: NOP   0;
NETWORK
TITLE =Step 9N1 - Power ON
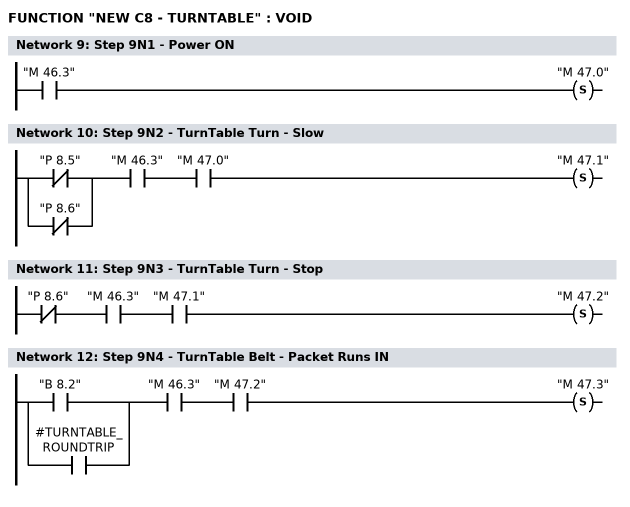

      A     "M 46.3";
      S     "M 47.0";
NETWORK
TITLE =Step 9N2 - TurnTable Turn - Slow

      A(    ;
      ON    "P 8.5";
      ON    "P 8.6";
      )     ;
      A     "M 46.3";
      A     "M 47.0";
      S     "M 47.1";
NETWORK
TITLE =Step 9N3 - TurnTable Turn - Stop

      AN    "P 8.6";
      A     "M 46.3";
      A     "M 47.1";
      S     "M 47.2";
NETWORK
TITLE =Step 9N4 - TurnTable Belt - Packet Runs IN

      A(    ;
      O     "B 8.2";
      O     #TURNTABLE_ROUNDTRIP;
      )     ;
      A     "M 46.3";
      A     "M 47.2";
      S     "M 47.3";
NETWORK
TITLE =Step 9N5 - TurnTable Belt 8 - Packet IN

      AN(   ;
      O     "B 8.2";
      O     #TURNTABLE_ROUNDTRIP;
      )     ;
      A     "M 46.3";
      A     "M 47.3";
      S     "M 47.4";
NETWORK
TITLE =TurnTable Belt Entry Jam Timeout
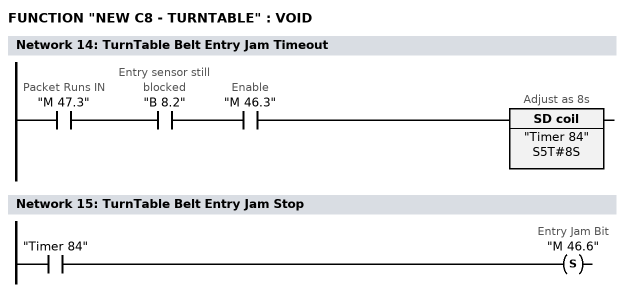

      A     "M 47.3"; // Packet Runs IN
      A     "B 8.2"; // Entry sensor still blocked
      A     "M 46.3"; // Enable
      L     S5T#8S; // Adjust as 8s
      SD    "Timer 84";
NETWORK
TITLE =TurnTable Belt Entry Jam Stop

      A     "Timer 84";
      S     "M 46.6"; // Entry Jam Bit
NETWORK
TITLE =Length Convertion - TurnTable Belt

      A     "M 31.4";
      FP    "FP 157.3";
      JNB   M317;
      L     "COLLATORS DB".PacketLength_C4;
      ITD   ;
      DTR   ;
      T     #PACKET_LENGTH;

      CALL "SCALER" (
           X                        := #PACKET_LENGTH,
           X1                       := 5.500000e+001,
           Y1                       := 2.000000e+003,
           X2                       := 1.600000e+002,
           Y2                       := 1.000000e+003,
           RET_VAL                  := #RUN_TIME);

      L     #RUN_TIME;
      RND   ;
      T     "MW 196";

M317: NOP   0;
NETWORK
TITLE =Time Convertion - TurnTable Belt
//- Packet Forward : - Run Time   (~1500mS)
//- Packet Reverse : - Run Time   (~300mS)
//950mm Packet : 1300 mS
//Collator 4 - 950 mm = 143 Count  6.6mm per pulse
//
//- Packet Inverting on TurnTable - Belt RunTime at Packet End: Always 300mS to
//Stay Close to REV Exit Side !
//
//- Packet Non-Inverting on TurnTable - Belt RunTime at Packet End: 500 to 1600mS
//(Depend on Packet Length) to get Close to FWD Exit Side !...
//
//404 Tube Limit 350 - 1050mm
      AN    "M 7.3";
      AN    "M 6.7";
      FP    "FP 157.6";
      JNB   END;
      L     "HMI_DB".CONV_8_POS_REV_mS; // Integer contains MILLISECOND seconds
      L     10;
      *I    ;
      ITD   ;
      T     #ZOOLOO;

      CALL "TIM_S5TI" (
           IN                       := #ZOOLOO,
           RET_VAL                  := "MW 234");

END:  NOP   0;
NETWORK
TITLE =TurnTable Belt  - Run Time FWD & REV  300mS
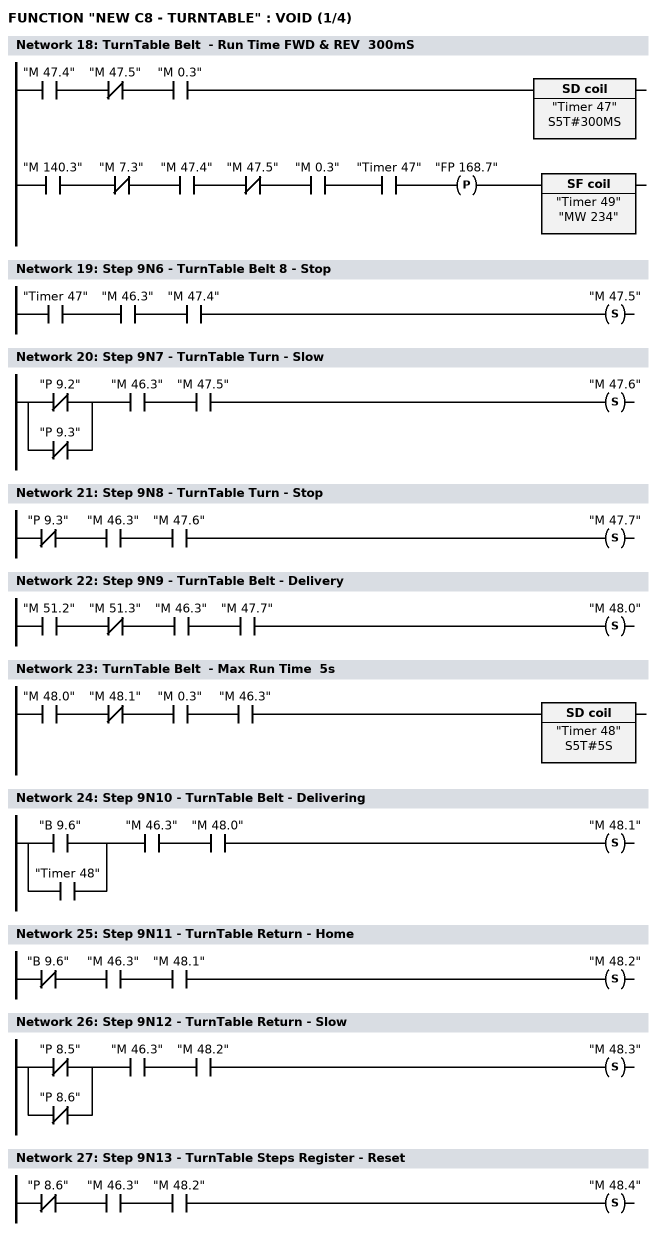

      A     "M 47.4";
      AN    "M 47.5";
      A     "M 0.3";
      L     S5T#300MS;
      SD    "Timer 47";
//;
      A     "M 140.3";
      AN    "M 7.3";
      A     "M 47.4";
      AN    "M 47.5";
      A     "M 0.3";
      A     "Timer 47";
      FP    "FP 168.7";
      L     "MW 234";
      SF    "Timer 49";
NETWORK
TITLE =Step 9N6 - TurnTable Belt 8 - Stop

      A     "Timer 47";
      A     "M 46.3";
      A     "M 47.4";
      S     "M 47.5";
NETWORK
TITLE =Step 9N7 - TurnTable Turn - Slow

      A(    ;
      ON    "P 9.2";
      ON    "P 9.3";
      )     ;
      A     "M 46.3";
      A     "M 47.5";
      S     "M 47.6";
NETWORK
TITLE =Step 9N8 - TurnTable Turn - Stop

      AN    "P 9.3";
      A     "M 46.3";
      A     "M 47.6";
      S     "M 47.7";
NETWORK
TITLE =Step 9N9 - TurnTable Belt - Delivery

      A     "M 51.2";
      AN    "M 51.3";
      A     "M 46.3";
      A     "M 47.7";
      S     "M 48.0";
NETWORK
TITLE =TurnTable Belt  - Max Run Time  5s

      A     "M 48.0";
      AN    "M 48.1";
      A     "M 0.3";
      A     "M 46.3";
      L     S5T#5S;
      SD    "Timer 48";
NETWORK
TITLE =Step 9N10 - TurnTable Belt - Delivering

      A(    ;
      O     "B 9.6";
      O     "Timer 48";
      )     ;
      A     "M 46.3";
      A     "M 48.0";
      S     "M 48.1";
NETWORK
TITLE =Step 9N11 - TurnTable Return - Home

      AN    "B 9.6";
      A     "M 46.3";
      A     "M 48.1";
      S     "M 48.2";
NETWORK
TITLE =Step 9N12 - TurnTable Return - Slow

      A(    ;
      ON    "P 8.5";
      ON    "P 8.6";
      )     ;
      A     "M 46.3";
      A     "M 48.2";
      S     "M 48.3";
NETWORK
TITLE =Step 9N13 - TurnTable Steps Register - Reset

      AN    "P 8.6";
      A     "M 46.3";
      A     "M 48.2";
      S     "M 48.4";
NETWORK
TITLE =Service Home Position Process - Position Home Test
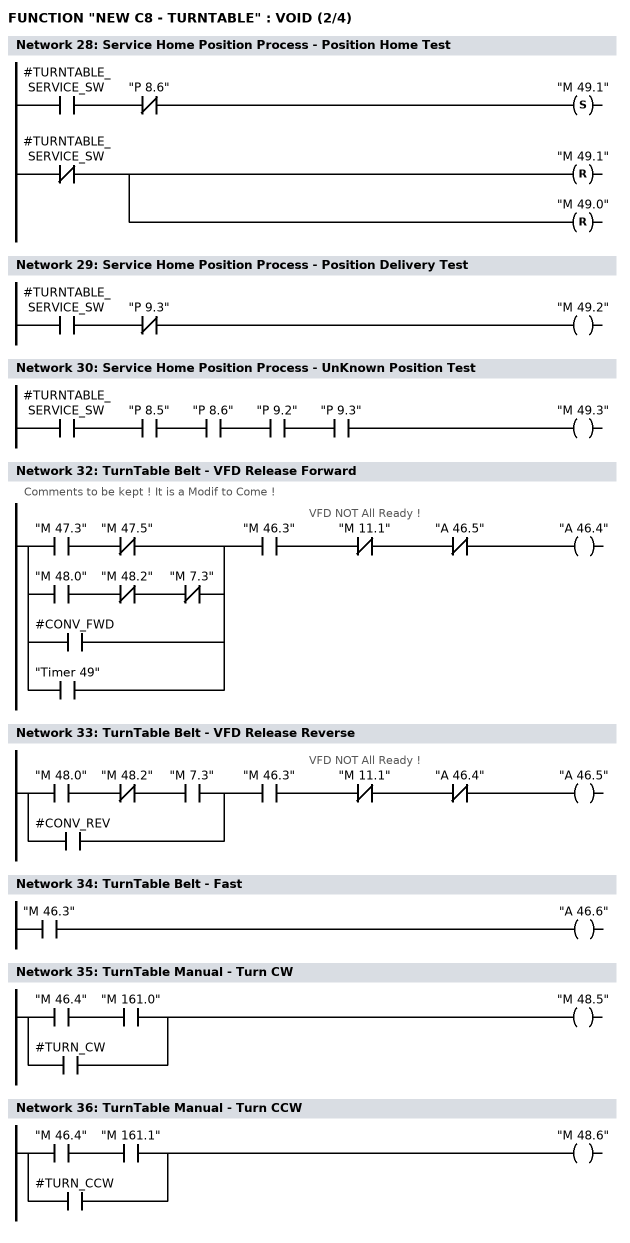

      A     #TURNTABLE_SERVICE_SW;
      AN    "P 8.6";
      S     "M 49.1";
//;
      AN    #TURNTABLE_SERVICE_SW;
      R     "M 49.1";
      R     "M 49.0";
NETWORK
TITLE =Service Home Position Process - Position Delivery Test

      A     #TURNTABLE_SERVICE_SW;
      AN    "P 9.3";
      =     "M 49.2";
NETWORK
TITLE =Service Home Position Process - UnKnown Position Test

      A     #TURNTABLE_SERVICE_SW;
      A     "P 8.5";
      A     "P 8.6";
      A     "P 9.2";
      A     "P 9.3";
      =     "M 49.3";
NETWORK
TITLE =Action from Steps Commands



NETWORK
TITLE =TurnTable Belt - VFD Release Forward
//Comments to be kept ! It is a Modif to Come !
      A(    ;
      A     "M 47.3";
      AN    "M 47.5";
      O     ;
      A     "M 48.0";
      AN    "M 48.2";
      AN    "M 7.3";
      )     ;
      O     #CONV_FWD;
      O     "Timer 49";
      A     "M 46.3";
      AN    "M 11.1"; // VFD NOT All Ready !
      AN    "A 46.5";
      =     "A 46.4";
NETWORK
TITLE =TurnTable Belt - VFD Release Reverse

      A(    ;
      A     "M 48.0";
      AN    "M 48.2";
      A     "M 7.3";
      O     #CONV_REV;
      )     ;
      A     "M 46.3";
      AN    "M 11.1"; // VFD NOT All Ready !
      AN    "A 46.4";
      =     "A 46.5";
NETWORK
TITLE =TurnTable Belt - Fast

      A     "M 46.3";
      =     "A 46.6";
NETWORK
TITLE =TurnTable Manual - Turn CW

      A     "M 46.4";
      A     "M 161.0";
      O     #TURN_CW;
      =     "M 48.5";
NETWORK
TITLE =TurnTable Manual - Turn CCW

      A     "M 46.4";
      A     "M 161.1";
      O     #TURN_CCW;
      =     "M 48.6";
NETWORK
TITLE =TurnTable Manual - Manual Mode Reset
